(* IEC 61131-3 sources: plc-iiot-stack/tests/POUs/FB_MqttCommands_Test, 18 files *)

(* ---- AcceptedStartWaitsForDeviceThenOk.method.decl.st ---- *)
// Start прошёл шлюз: stCmd, ответа нет до обработки устройством, затем ok.
METHOD PRIVATE AcceptedStartWaitsForDeviceThenOk
VAR_INST
    fbFake : FB_MqttClientFake;
    fbCmd : FB_MqttCommands;
    aRules : ARRAY[1..4] OF ST_IiotCmdRule;
END_VAR

(* ---- DeviceRejectedCarriesCmdResult.method.decl.st ---- *)
// Устройство отказало — device_rejected и cmd_result по E_CmdResult.
METHOD PRIVATE DeviceRejectedCarriesCmdResult
VAR_INST
    fbFake : FB_MqttClientFake;
    fbCmd : FB_MqttCommands;
    aRules : ARRAY[1..4] OF ST_IiotCmdRule;
END_VAR

(* ---- DeviceSilenceIsTimeout.method.decl.st ---- *)
// Устройство не обработало команду за 3 с — timeout; новое сообщение ждёт.
METHOD PRIVATE DeviceSilenceIsTimeout
VAR_INST
    fbFake : FB_MqttClientFake;
    fbCmd : FB_MqttCommands;
    aRules : ARRAY[1..4] OF ST_IiotCmdRule;
END_VAR

(* ---- DropsWithoutAckWhenNoCmdId.method.decl.st ---- *)
// Не своя станция, не JSON, нет или неверный cmd_id, обрезано — без ответа.
METHOD PRIVATE DropsWithoutAckWhenNoCmdId
VAR_INST
    fbFake : FB_MqttClientFake;
    fbCmd : FB_MqttCommands;
    aRules : ARRAY[1..4] OF ST_IiotCmdRule;
END_VAR

(* ---- MissingArmMeansTimeout.method.decl.st ---- *)
// Команда прошла шлюз, но Arm() не вызван — ответ timeout в следующем вызове.
METHOD PRIVATE MissingArmMeansTimeout
VAR_INST
    fbFake : FB_MqttClientFake;
    fbCmd : FB_MqttCommands;
    aRules : ARRAY[1..4] OF ST_IiotCmdRule;
END_VAR

(* ---- RateLimitTenPerTenSeconds.method.decl.st ---- *)
// Не больше 10 команд за 10 с — rate_limited; после окна — снова принимаются.
METHOD PRIVATE RateLimitTenPerTenSeconds
VAR_INST
    fbFake : FB_MqttClientFake;
    fbCmd : FB_MqttCommands;
    aRules : ARRAY[1..4] OF ST_IiotCmdRule;
END_VAR

(* ---- RejectsDuplicateIncludingRejectedIds.method.decl.st ---- *)
// Повтор cmd_id среди последних 16 (и отклонённых тоже) — duplicate.
METHOD PRIVATE RejectsDuplicateIncludingRejectedIds
VAR_INST
    fbFake : FB_MqttClientFake;
    fbCmd : FB_MqttCommands;
    aRules : ARRAY[1..4] OF ST_IiotCmdRule;
END_VAR

(* ---- RejectsExpired.method.decl.st ---- *)
// ts дальше 30 с от часов ПЛК (в прошлое или будущее) или часов нет — expired.
METHOD PRIVATE RejectsExpired
VAR_INST
    fbFake : FB_MqttClientFake;
    fbCmd : FB_MqttCommands;
    aRules : ARRAY[1..4] OF ST_IiotCmdRule;
END_VAR

(* ---- RejectsInvalidPayloads.method.decl.st ---- *)
// Не по command.schema.json — invalid_payload: лишние поля, ts, origin, command, value.
METHOD PRIVATE RejectsInvalidPayloads
VAR_INST
    fbFake : FB_MqttClientFake;
    fbCmd : FB_MqttCommands;
    aRules : ARRAY[1..4] OF ST_IiotCmdRule;
END_VAR

(* ---- RejectsNotWhitelisted.method.decl.st ---- *)
// Пары (устройство, команда) нет в белом списке — not_whitelisted.
METHOD PRIVATE RejectsNotWhitelisted
VAR_INST
    fbFake : FB_MqttClientFake;
    fbCmd : FB_MqttCommands;
    aRules : ARRAY[1..4] OF ST_IiotCmdRule;
END_VAR

(* ---- RejectsOutOfRange.method.decl.st ---- *)
// SpeedSp вне 0..100 % — out_of_range.
METHOD PRIVATE RejectsOutOfRange
VAR_INST
    fbFake : FB_MqttClientFake;
    fbCmd : FB_MqttCommands;
    aRules : ARRAY[1..4] OF ST_IiotCmdRule;
END_VAR

(* ---- RejectsRetainedCommand.method.decl.st ---- *)
// Команда с флагом retain — retained.
METHOD PRIVATE RejectsRetainedCommand
VAR_INST
    fbFake : FB_MqttClientFake;
    fbCmd : FB_MqttCommands;
    aRules : ARRAY[1..4] OF ST_IiotCmdRule;
END_VAR

(* ---- RejectsUnsupportedVersionAndTopicMismatch.method.decl.st ---- *)
// schema_version 2.0 — unsupported_version; команда не та, что в топике.
METHOD PRIVATE RejectsUnsupportedVersionAndTopicMismatch
VAR_INST
    fbFake : FB_MqttClientFake;
    fbCmd : FB_MqttCommands;
    aRules : ARRAY[1..4] OF ST_IiotCmdRule;
END_VAR

(* ---- Run.method.decl.st ---- *)
// Поставить сообщение в очередь (sTopic пусто — без сообщения) и вызвать FB_MqttCommands.
METHOD PRIVATE Run
VAR_IN_OUT
    fbClient : FB_MqttClientFake;
    fbCommands : FB_MqttCommands;
    aRuleTable : ARRAY[*] OF ST_IiotCmdRule;
END_VAR
VAR_INPUT
    sTopic : STRING(GVL_Const.MQTT_TOPIC_LEN) := '';
    sPayload : STRING(GVL_Const.MQTT_CMD_PAYLOAD_LEN) := '';
    xRetainedIn : BOOL := FALSE;
    ltAt : LTIME := LTIME#1H;
    uliNow_ms : ULINT := 1792137600250;
    uiSeq : UINT := 0;
    iResult : INT := 0;
END_VAR

(* ---- Run.method.impl.st ---- *)
IF LEN(sTopic) > 0 THEN
    fbClient.Inject(sTopic := sTopic, sPayload := sPayload, xTruncated := FALSE, xRetained := xRetainedIn);
END_IF
fbCommands(xEnable := TRUE, itfClient := fbClient, ltNow := ltAt, uliTs_ms := uliNow_ms,
           sTopicPrefix := 'vodokanal/kns1/station', uiDevSeq := uiSeq, iDevResult := iResult, aRules := aRuleTable);

(* ---- Setup.method.decl.st ---- *)
// Белый список: P101 Start, SpeedSp (0..100 %), Ack; LT101 Ack. Связь есть.
METHOD PRIVATE Setup
VAR_IN_OUT
    fbClient : FB_MqttClientFake;
    aRuleTable : ARRAY[1..4] OF ST_IiotCmdRule;
END_VAR

(* ---- SpeedSetpointIsOkAfterWrite.method.decl.st ---- *)
// SpeedSp: ok сразу после записи (ФБ устройства значения не квитирует); границы 0 и 100.
METHOD PRIVATE SpeedSetpointIsOkAfterWrite
VAR_INST
    fbFake : FB_MqttClientFake;
    fbCmd : FB_MqttCommands;
    aRules : ARRAY[1..4] OF ST_IiotCmdRule;
END_VAR

(* ---- SubscribesToCommandTopicsAndResubscribes.method.decl.st ---- *)
// Подписка <site>/<area>/<unit>/+/cmd/+ с QoS 1; заново после переподключения.
METHOD PRIVATE SubscribesToCommandTopicsAndResubscribes
VAR_INST
    fbFake : FB_MqttClientFake;
    fbCmd : FB_MqttCommands;
    aRules : ARRAY[1..4] OF ST_IiotCmdRule;
END_VAR
